{attribute 'linkalways'}
{attribute 'no_explicit_call' := 'Use the methods of this class'}
{attribute 'enable_dynamic_creation'}
FUNCTION_BLOCK Lidar_Simulated IMPLEMENTS I_Lidar
VAR
	notConnectedError : HardwareError := (isActive := TRUE, id := Constants.SIMULATOR_NOT_CONNECTED_ERROR_ID, text := 'Simulatoren er ikke tilkoblet');
	link : REFERENCE TO SimulatorLink;
	_isRunning : BOOL;
	lastSequence : UDINT;
END_VAR

METHOD FB_init : BOOL
VAR_INPUT
	bInitRetains : BOOL;
	bInCopyCode : BOOL;
	simulator : REFERENCE TO SimulatorLink;
END_VAR
link REF= simulator;
END_METHOD

METHOD Start
_isRunning := TRUE;
lastSequence := SimulatorIo.scan.sequence;
END_METHOD

METHOD Stop
_isRunning := FALSE;
END_METHOD

METHOD TryGetScan : BOOL
VAR_INPUT
	scan : REFERENCE TO LaserScan;
END_VAR
IF NOT _isRunning OR_ELSE SimulatorIo.scan.sequence = lastSequence THEN
	RETURN;
END_IF
lastSequence := SimulatorIo.scan.sequence;
scan := SimulatorIo.scan;
TryGetScan := TRUE;
END_METHOD

PROPERTY IsRunning : BOOL
GET
IsRunning := _isRunning;
END_GET
END_PROPERTY

PROPERTY Error : HardwareError
GET
IF NOT __ISVALIDREF(link) OR_ELSE NOT link.IsConnected THEN
	Error := notConnectedError;
END_IF
END_GET
END_PROPERTY

END_FUNCTION_BLOCK

(* stored: Version 1.1.0.1, ProductVersion 3.1.4026.12
   POU Lidar_Simulated: Id {f8a143f8-acdc-5460-933b-52bfb9af5326}, SpecialFunc None
   Method FB_init: Id {fc740cba-7289-561c-b90d-5fd3eff46435}
   Method Start: Id {03fce770-f4df-52ae-8699-2b3d6feada58}
   Method Stop: Id {dcbf6750-aa7a-585e-868d-049504cf92a4}
   Method TryGetScan: Id {23df3983-3889-5989-b13a-c98300787fbf}
   Property IsRunning: Id {c9b9c1e0-5c86-51ec-a8a5-3edfe93d73b5}
   Get Get: Id {1f9915ee-0f5e-5956-8166-a1df040b8fe4}
   Property Error: Id {ef917698-682e-568a-9815-494f41f67a64}
   Get Get: Id {fad89dfc-b12c-549c-9702-76cce736f1fa} *)
